// TIA Portal project "sorting by height" (V17)
// Vorlageprojekt für das Buch mit Zielsystem S7-1200

(* hardware
DEVICE "S7-1200-Station_1"  S7-1200 Station
   slot 0: "Baugruppenträger_0"  Rack  V1.0
   slot 1: "PLC_1"  CPU 1211C DC/DC/DC  6ES7 211-1AE40-0XB0  V4.1
*)

// ===== PLC "PLC_1"  CPU 1211C DC/DC/DC =====

VAR_GLOBAL   // PLC tag table "sorting"
   "start" AT %I0.0 : Bool;
   "stop" AT %I0.1 : Bool;
   "low_sensor" AT %I0.3 : Bool;
   "high_sensor" AT %I0.4 : Bool;
   "loaded_sensor" AT %I0.5 : Bool;
   "right_entry_sensor" AT %I0.6 : Bool;
   "left_entry_sensor" AT %I0.7 : Bool;
   "trans_right" AT %Q0.0 : Bool;
   "trans_left" AT %Q0.1 : Bool;
   "conv_right" AT %Q0.2 : Bool;
   "conv_left" AT %Q0.3 : Bool;
   "pallet_sensor" AT %I1.0 : Bool;
   "load_conveyor" AT %Q0.4 : Bool;
   "right_exit_sensor" AT %I1.1 : Bool;
   "left_exit_sensor" AT %I1.2 : Bool;
   "coveyor_entry" AT %Q0.5 : Bool;
   "Reset" AT %I1.3 : Bool;
   "emergency_stop" AT %I0.2 : Bool;
   "counter" AT %QW30 : Word;
   "Clock_Byte" AT %MB100 : Byte;
   "Clock_10Hz" AT %M100.0 : Bool;
   "Clock_5Hz" AT %M100.1 : Bool;
   "Clock_2.5Hz" AT %M100.2 : Bool;
   "Clock_2Hz" AT %M100.3 : Bool;
   "Clock_1.25Hz" AT %M100.4 : Bool;
   "Clock_1Hz" AT %M100.5 : Bool;
   "Clock_0.625Hz" AT %M100.6 : Bool;
   "Clock_0.5Hz" AT %M100.7 : Bool;
   "Start_light" AT %Q0.6 : Bool;
   "Stop_light" AT %Q0.7 : Bool;
   "Reset_light" AT %Q1.0 : Bool;
   "System_Byte" AT %MB1 : Byte;
   "FirstScan" AT %M1.0 : Bool;
   "DiagStatusUpdate" AT %M1.1 : Bool;
   "AlwaysTRUE" AT %M1.2 : Bool;
   "AlwaysFALSE" AT %M1.3 : Bool;
END_VAR

DATA_BLOCK "DB"   // DB1
{ S7_Optimized_Access := 'TRUE' }
VERSION : 0.1
   VAR
      Infeed_Conveyor : Bool;
      RIght_Conveyor : Bool;
      Left_Conveyor : Bool;
      load_coveyor : Bool;
      high_active : Bool;
      low_active : Bool;
      right_entry : Bool;
      left_entry : Bool;
      left_exit : Bool;
      right_exit : Bool;
      system_on : Bool;
      p_trigger : Bool;
   END_VAR
BEGIN
END_DATA_BLOCK

// folder: System blocks/Program resources

DATA_BLOCK "Box_count"   // DB2
{ S7_Optimized_Access := 'TRUE' }
AUTHOR : Simatic
FAMILY : IEC
NAME : CNTR
VERSION : 1.0
// stored: InstanceOfName IEC_COUNTER
"IEC_COUNTER"
BEGIN
END_DATA_BLOCK

DATA_BLOCK "trans_right_delay"   // DB3
{ S7_Optimized_Access := 'TRUE' }
AUTHOR : Simatic
FAMILY : IEC
NAME : IEC_TMR
VERSION : 1.0
// stored: InstanceOfName IEC_TIMER
"IEC_TIMER"
BEGIN
END_DATA_BLOCK

DATA_BLOCK "trans_left_delay"   // DB4
{ S7_Optimized_Access := 'TRUE' }
AUTHOR : Simatic
FAMILY : IEC
NAME : IEC_TMR
VERSION : 1.0
// stored: InstanceOfName IEC_TIMER
"IEC_TIMER"
BEGIN
END_DATA_BLOCK

// folder: (top level)

FUNCTION "State handler" : Void   // FC1, LAD
{ S7_Optimized_Access := 'TRUE' }
VERSION : 0.1
BEGIN

REGION Network 1: fault safe
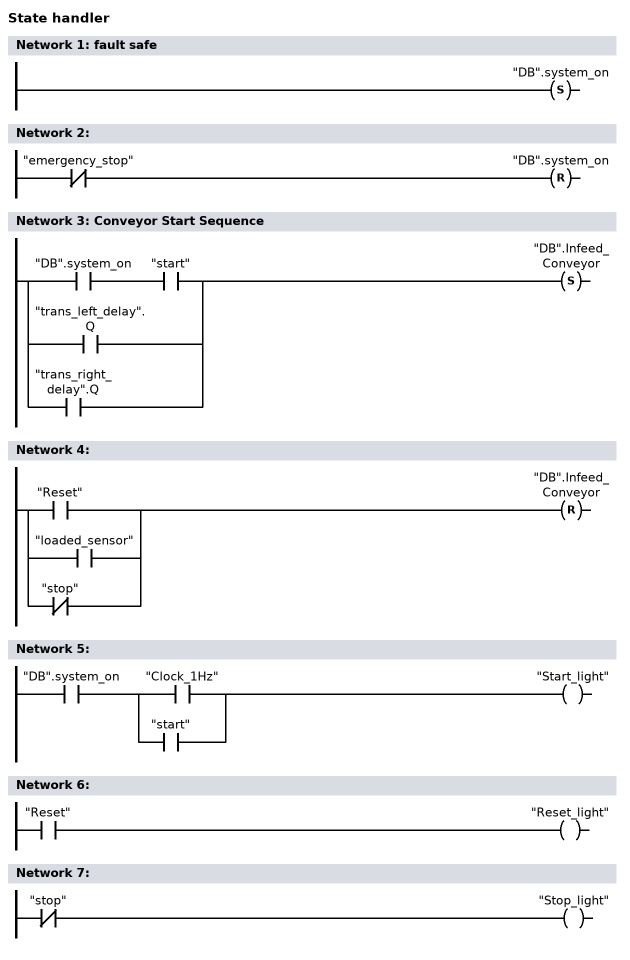
   RUNG wire#powerrail
      S_Coil( "DB".system_on )
   END_RUNG
   // the same network as SCL:
   "DB".system_on := TRUE;
END_REGION

REGION Network 2
   RUNG wire#powerrail
      I_Contact( "emergency_stop" )
      R_Coil( "DB".system_on )
   END_RUNG
   // the same network as SCL:
   IF NOT "emergency_stop" THEN "DB".system_on := FALSE; END_IF;
END_REGION

REGION Network 3: Conveyor Start Sequence
   RUNG wire#powerrail
      Contact( "DB".system_on )
      Contact( "start" )
      wire#w1
      S_Coil( "DB".Infeed_Conveyor )
   END_RUNG
   RUNG wire#powerrail
      Contact( "trans_left_delay".Q )
   END_RUNG wire#w1
   RUNG wire#powerrail
      Contact( "trans_right_delay".Q )
   END_RUNG wire#w1
   // the same network as SCL:
   IF ("DB".system_on AND "start") OR "trans_left_delay".Q OR "trans_right_delay".Q THEN
       "DB".Infeed_Conveyor := TRUE;
   END_IF;
END_REGION

REGION Network 4
   RUNG wire#powerrail
      Contact( "Reset" )
      wire#w1
      R_Coil( "DB".Infeed_Conveyor )
   END_RUNG
   RUNG wire#powerrail
      Contact( "loaded_sensor" )
   END_RUNG wire#w1
   RUNG wire#powerrail
      I_Contact( "stop" )
   END_RUNG wire#w1
   // the same network as SCL:
   IF "Reset" OR "loaded_sensor" OR NOT "stop" THEN "DB".Infeed_Conveyor := FALSE; END_IF;
END_REGION

REGION Network 5
   RUNG wire#powerrail
      Contact( "DB".system_on )
      wire#w1
      Contact( "Clock_1Hz" )
      wire#w2
      Coil( "Start_light" )
   END_RUNG
   RUNG wire#w1
      Contact( "start" )
   END_RUNG wire#w2
   // the same network as SCL:
   "Start_light" := "DB".system_on AND ("Clock_1Hz" OR "start");
END_REGION

REGION Network 6
   RUNG wire#powerrail
      Contact( "Reset" )
      Coil( "Reset_light" )
   END_RUNG
   // the same network as SCL:
   "Reset_light" := "Reset";
END_REGION

REGION Network 7
   RUNG wire#powerrail
      I_Contact( "stop" )
      Coil( "Stop_light" )
   END_RUNG
   // the same network as SCL:
   "Stop_light" := NOT "stop";
END_REGION
END_FUNCTION

FUNCTION "MHJ-PLC-Lab-Function-S71200" : Void   // FC9000, SCL
{ S7_Optimized_Access := 'TRUE' }
VERSION : 0.1
   VAR_TEMP
      rdTimeReturn : Int;
      outputTime : DTL;
      SyncVal : Byte;
      forVal : Int;
      forVal_2 : Int;
      Value : Byte;
   END_VAR
   VAR CONSTANT
      CompVal : Byte := 16#34;
      Value_01 : Byte := 16#11;
      Value_01_DW : DWord := 16#A165_D992;
      Value_02_DW : DWord := 16#58BE_4401;
   END_VAR
BEGIN

   #Value:=PEEK(area := 16#82,
        dbNumber := 0,
        byteOffset := 511);
   #Value := #Value + 1;

   POKE(area := 16#82,
        dbNumber := 0,
        byteOffset := 511,
        value := #Value);

   POKE(area:=16#81,
        dbNumber:=0,
        byteOffset:=1016,
        value:=#Value_01_DW);
   POKE(area := 16#81,
        dbNumber := 0,
        byteOffset := 1020,
        value := #Value_02_DW);

   POKE(area := 16#81,
        dbNumber := 0,
        byteOffset := 511,
        value := B#16#00);

   FOR #forVal := 0 TO 120 DO
       FOR #forVal_2:=0 TO 10 DO
           #rdTimeReturn:=RD_SYS_T(#outputTime);
           #rdTimeReturn := WR_SYS_T(#outputTime);
           #rdTimeReturn := RD_SYS_T(#outputTime);
           #rdTimeReturn := WR_SYS_T(#outputTime);
       END_FOR;
       #SyncVal:= PEEK(area := 16#81,
                      dbNumber := 0,
                      byteOffset := 511);
       IF #SyncVal = #CompVal THEN
          GOTO M_1;
       END_IF;
   END_FOR;
   RETURN;

   M_1:
   POKE(area := 16#81,
        dbNumber := 0,
        byteOffset := 511,
        value := B#16#0);
END_FUNCTION

ORGANIZATION_BLOCK "Main"   // OB1, LAD, ProgramCycle
TITLE = "Main Program Sweep (Cycle)"
{ S7_Optimized_Access := 'TRUE' }
VERSION : 0.1
   VAR_INPUT
      Initial_Call : Bool;   // Initial call of this OB
      Remanence : Bool;   // =True, if remanent data are available
   END_VAR
   VAR_TEMP   // added for the SCL form of the ladder/FBD networks
      _w1 : Bool;
   END_VAR
BEGIN

REGION Network 1
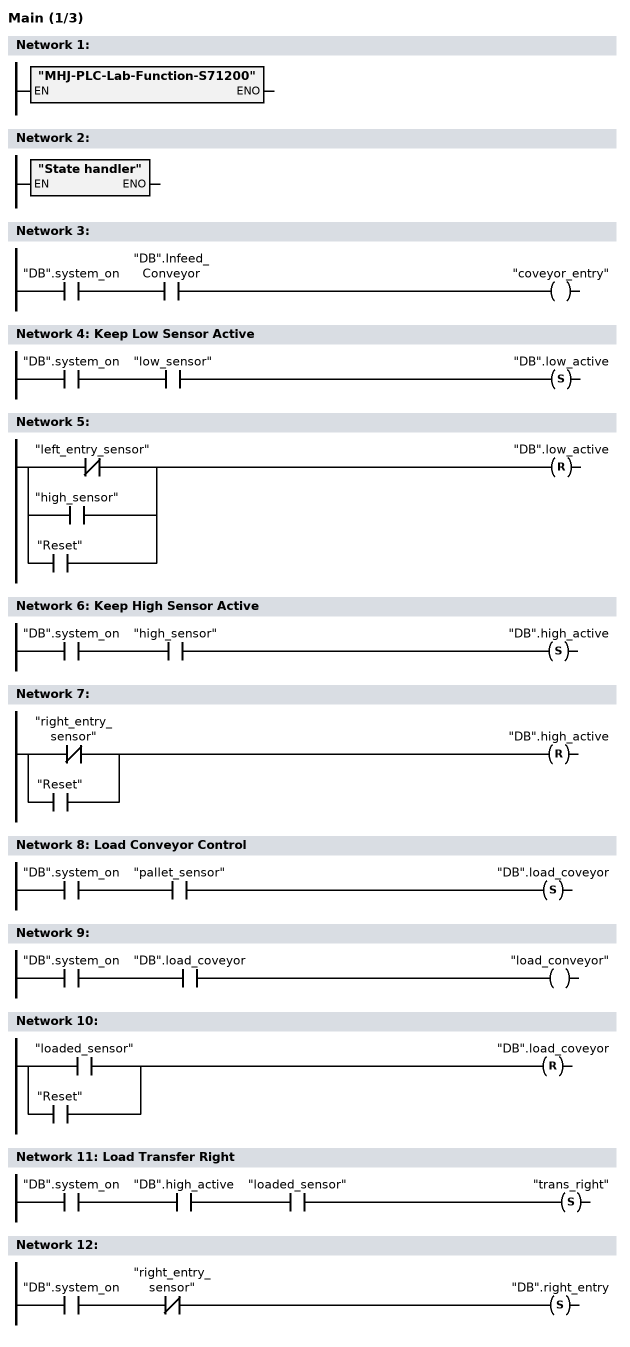
   RUNG wire#powerrail
      "MHJ-PLC-Lab-Function-S71200"()
   END_RUNG
   // the same network as SCL:
   "MHJ-PLC-Lab-Function-S71200"();
END_REGION

REGION Network 2
   RUNG wire#powerrail
      "State handler"()
   END_RUNG
   // the same network as SCL:
   "State handler"();
END_REGION

REGION Network 3
   RUNG wire#powerrail
      Contact( "DB".system_on )
      Contact( "DB".Infeed_Conveyor )
      Coil( "coveyor_entry" )
   END_RUNG
   // the same network as SCL:
   "coveyor_entry" := "DB".system_on AND "DB".Infeed_Conveyor;
END_REGION

REGION Network 4: Keep Low Sensor Active
   RUNG wire#powerrail
      Contact( "DB".system_on )
      Contact( "low_sensor" )
      S_Coil( "DB".low_active )
   END_RUNG
   // the same network as SCL:
   IF "DB".system_on AND "low_sensor" THEN "DB".low_active := TRUE; END_IF;
END_REGION

REGION Network 5
   RUNG wire#powerrail
      I_Contact( "left_entry_sensor" )
      wire#w1
      R_Coil( "DB".low_active )
   END_RUNG
   RUNG wire#powerrail
      Contact( "high_sensor" )
   END_RUNG wire#w1
   RUNG wire#powerrail
      Contact( "Reset" )
   END_RUNG wire#w1
   // the same network as SCL:
   IF NOT "left_entry_sensor" OR "high_sensor" OR "Reset" THEN "DB".low_active := FALSE; END_IF;
END_REGION

REGION Network 6: Keep High Sensor Active
   RUNG wire#powerrail
      Contact( "DB".system_on )
      Contact( "high_sensor" )
      S_Coil( "DB".high_active )
   END_RUNG
   // the same network as SCL:
   IF "DB".system_on AND "high_sensor" THEN "DB".high_active := TRUE; END_IF;
END_REGION

REGION Network 7
   RUNG wire#powerrail
      I_Contact( "right_entry_sensor" )
      wire#w1
      R_Coil( "DB".high_active )
   END_RUNG
   RUNG wire#powerrail
      Contact( "Reset" )
   END_RUNG wire#w1
   // the same network as SCL:
   IF NOT "right_entry_sensor" OR "Reset" THEN "DB".high_active := FALSE; END_IF;
END_REGION

REGION Network 8: Load Conveyor Control
   RUNG wire#powerrail
      Contact( "DB".system_on )
      Contact( "pallet_sensor" )
      S_Coil( "DB".load_coveyor )
   END_RUNG
   // the same network as SCL:
   IF "DB".system_on AND "pallet_sensor" THEN "DB".load_coveyor := TRUE; END_IF;
END_REGION

REGION Network 9
   RUNG wire#powerrail
      Contact( "DB".system_on )
      Contact( "DB".load_coveyor )
      Coil( "load_conveyor" )
   END_RUNG
   // the same network as SCL:
   "load_conveyor" := "DB".system_on AND "DB".load_coveyor;
END_REGION

REGION Network 10
   RUNG wire#powerrail
      Contact( "loaded_sensor" )
      wire#w1
      R_Coil( "DB".load_coveyor )
   END_RUNG
   RUNG wire#powerrail
      Contact( "Reset" )
   END_RUNG wire#w1
   // the same network as SCL:
   IF "loaded_sensor" OR "Reset" THEN "DB".load_coveyor := FALSE; END_IF;
END_REGION

REGION Network 11: Load Transfer Right
   RUNG wire#powerrail
      Contact( "DB".system_on )
      Contact( "DB".high_active )
      Contact( "loaded_sensor" )
      S_Coil( "trans_right" )
   END_RUNG
   // the same network as SCL:
   IF "DB".system_on AND "DB".high_active AND "loaded_sensor" THEN "trans_right" := TRUE; END_IF;
END_REGION

REGION Network 12
   RUNG wire#powerrail
      Contact( "DB".system_on )
      I_Contact( "right_entry_sensor" )
      S_Coil( "DB".right_entry )
   END_RUNG
   // the same network as SCL:
   IF "DB".system_on AND NOT "right_entry_sensor" THEN "DB".right_entry := TRUE; END_IF;
END_REGION

REGION Network 13
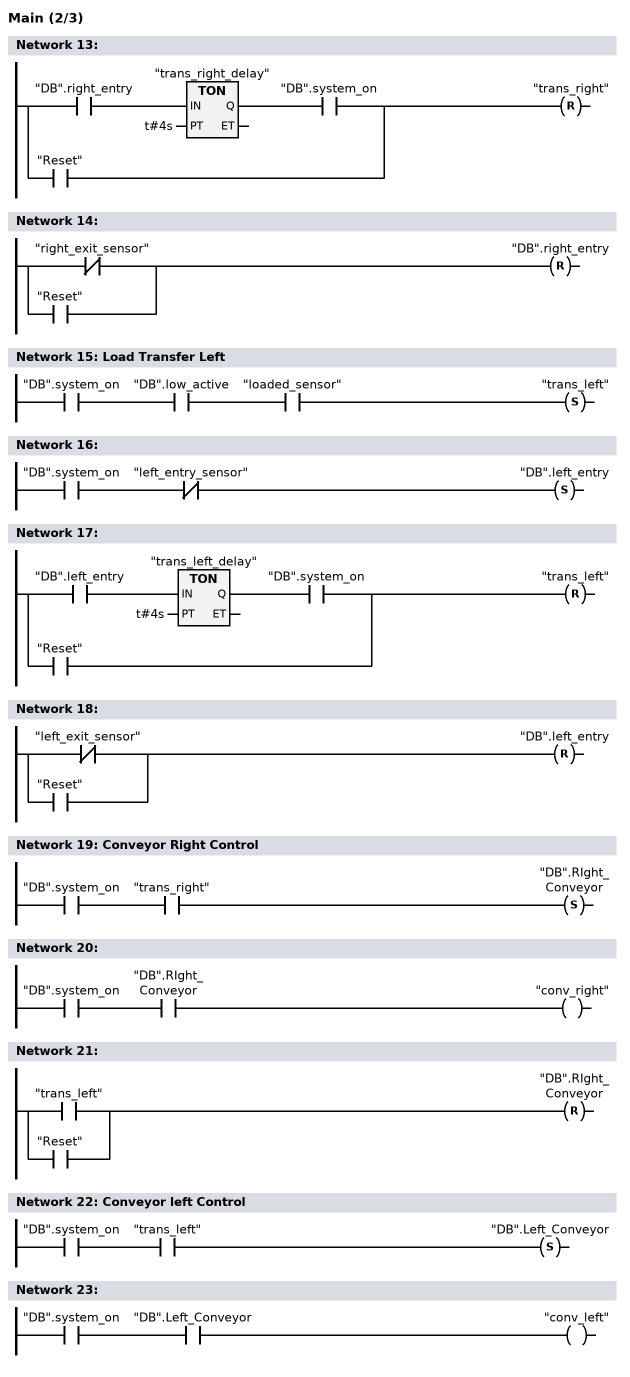
   "trans_right_delay".TON(IN := "DB".right_entry, PT := t#4s);
   IF ("trans_right_delay".Q AND "DB".system_on) OR "Reset" THEN "trans_right" := FALSE; END_IF;
END_REGION

REGION Network 14
   RUNG wire#powerrail
      I_Contact( "right_exit_sensor" )
      wire#w1
      R_Coil( "DB".right_entry )
   END_RUNG
   RUNG wire#powerrail
      Contact( "Reset" )
   END_RUNG wire#w1
   // the same network as SCL:
   IF NOT "right_exit_sensor" OR "Reset" THEN "DB".right_entry := FALSE; END_IF;
END_REGION

REGION Network 15: Load Transfer Left
   RUNG wire#powerrail
      Contact( "DB".system_on )
      Contact( "DB".low_active )
      Contact( "loaded_sensor" )
      S_Coil( "trans_left" )
   END_RUNG
   // the same network as SCL:
   IF "DB".system_on AND "DB".low_active AND "loaded_sensor" THEN "trans_left" := TRUE; END_IF;
END_REGION

REGION Network 16
   RUNG wire#powerrail
      Contact( "DB".system_on )
      I_Contact( "left_entry_sensor" )
      S_Coil( "DB".left_entry )
   END_RUNG
   // the same network as SCL:
   IF "DB".system_on AND NOT "left_entry_sensor" THEN "DB".left_entry := TRUE; END_IF;
END_REGION

REGION Network 17
   "trans_left_delay".TON(IN := "DB".left_entry, PT := t#4s);
   IF ("trans_left_delay".Q AND "DB".system_on) OR "Reset" THEN "trans_left" := FALSE; END_IF;
END_REGION

REGION Network 18
   RUNG wire#powerrail
      I_Contact( "left_exit_sensor" )
      wire#w1
      R_Coil( "DB".left_entry )
   END_RUNG
   RUNG wire#powerrail
      Contact( "Reset" )
   END_RUNG wire#w1
   // the same network as SCL:
   IF NOT "left_exit_sensor" OR "Reset" THEN "DB".left_entry := FALSE; END_IF;
END_REGION

REGION Network 19: Conveyor Right Control
   RUNG wire#powerrail
      Contact( "DB".system_on )
      Contact( "trans_right" )
      S_Coil( "DB".RIght_Conveyor )
   END_RUNG
   // the same network as SCL:
   IF "DB".system_on AND "trans_right" THEN "DB".RIght_Conveyor := TRUE; END_IF;
END_REGION

REGION Network 20
   RUNG wire#powerrail
      Contact( "DB".system_on )
      Contact( "DB".RIght_Conveyor )
      Coil( "conv_right" )
   END_RUNG
   // the same network as SCL:
   "conv_right" := "DB".system_on AND "DB".RIght_Conveyor;
END_REGION

REGION Network 21
   RUNG wire#powerrail
      Contact( "trans_left" )
      wire#w1
      R_Coil( "DB".RIght_Conveyor )
   END_RUNG
   RUNG wire#powerrail
      Contact( "Reset" )
   END_RUNG wire#w1
   // the same network as SCL:
   IF "trans_left" OR "Reset" THEN "DB".RIght_Conveyor := FALSE; END_IF;
END_REGION

REGION Network 22: Conveyor left Control
   RUNG wire#powerrail
      Contact( "DB".system_on )
      Contact( "trans_left" )
      S_Coil( "DB".Left_Conveyor )
   END_RUNG
   // the same network as SCL:
   IF "DB".system_on AND "trans_left" THEN "DB".Left_Conveyor := TRUE; END_IF;
END_REGION

REGION Network 23
   RUNG wire#powerrail
      Contact( "DB".system_on )
      Contact( "DB".Left_Conveyor )
      Coil( "conv_left" )
   END_RUNG
   // the same network as SCL:
   "conv_left" := "DB".system_on AND "DB".Left_Conveyor;
END_REGION

REGION Network 24
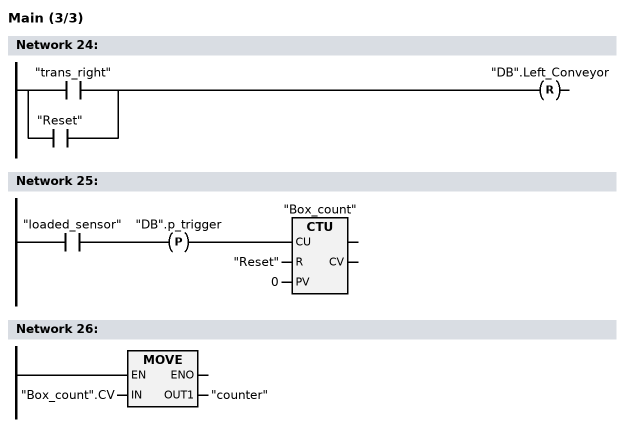
   RUNG wire#powerrail
      Contact( "trans_right" )
      wire#w1
      R_Coil( "DB".Left_Conveyor )
   END_RUNG
   RUNG wire#powerrail
      Contact( "Reset" )
   END_RUNG wire#w1
   // the same network as SCL:
   IF "trans_right" OR "Reset" THEN "DB".Left_Conveyor := FALSE; END_IF;
END_REGION

REGION Network 25
   #_w1 := "loaded_sensor" AND NOT "DB".p_trigger;   // rising edge
   "DB".p_trigger := "loaded_sensor";
   "Box_count".CTU(CU := #_w1, R := "Reset", PV := 0);
END_REGION

REGION Network 26
   RUNG wire#powerrail
      Move(in := "Box_count".CV, out1 => "counter")
   END_RUNG
   // the same network as SCL:
   "counter" := "Box_count".CV;
END_REGION
END_ORGANIZATION_BLOCK